FUNCTION VC_GetBool : BOOL
// Reads Bool (1 byte, little-endian) from Buf[Pos] and advances Pos.
VAR_IN_OUT
    Buf   : ARRAY[*] OF BYTE;
    Pos   : UDINT;
END_VAR
VAR
    nByte : BYTE;
END_VAR

nByte := 0;
VC_GetRaw(Buf := Buf, Pos := Pos, pDst := ADR(nByte), Size := 1);
VC_GetBool := (nByte <> 0);

END_FUNCTION

(* stored: Version 1.1.0.1, ProductVersion 3.1.4024.12
   POU VC_GetBool: Id {da520ad8-6b3e-4838-aea7-20d7e4599c1d}, SpecialFunc None *)
